// TIA Portal V21 export
// export: Created 2026-10-23T20:42:49.2153174Z, ExportSetting WithDefaults, DisplayName Totally Integrated Automation Portal, DisplayVersion V21 Update 1, DisplayName SINAMICS Startdrive Advanced, DisplayVersion V21 HF2, DisplayName SINAMICS Startdrive G110M, G120, G120C, G120D, G120P, G115D, DisplayVersion V21 HF2, DisplayName SINAMICS Startdrive G130, G150, S120, S150, G200, G220, S200, S210, S220, Innomotics MVD, DisplayVersion V21 HF2, DisplayName STEP 7 Professional, DisplayVersion V21 Update 1, DisplayName STEP 7 Safety, DisplayVersion V21, DisplayName Tech WebApplication, DisplayVersion V21, DisplayName WinCC Basic/Comfort/Advanced, DisplayVersion V21 Update 1, DisplayName WinCC Unified, DisplayVersion V21 Update 1
FUNCTION_BLOCK "FB_Mixed"   // FB9, LAD
TITLE = KOP-Baustein mit SCL-Netzwerk / LAD block with an SCL network
{ S7_Optimized_Access := 'TRUE' }
VERSION : 0.1
// stored: AutoNumber true, IsIECCheckEnabled false, IsRetainMemResEnabled false, MemoryReserve 100, SetENOAutomatically false, UDAEnableTagReadback false
   VAR_INPUT
      Start : Bool;   // Startbefehl / Start command
      RawValue : Int;   // Rohwert / Raw value
   END_VAR
   VAR_OUTPUT
      Running : Bool;   // Läuft / Running
      Scaled : Real;   // Skalierter Wert / Scaled value
      AboveLimit : Bool;   // Läuft und über dem Grenzwert / Running and above the limit
   END_VAR
   VAR
      Factor : Real := 2.5;   // Skalierungsfaktor / Scaling factor
      Limit : Real := 100.0;   // Grenzwert / Limit
      IsAbove : Bool;   // Skalierter Wert über dem Grenzwert / Scaled value above the limit
   END_VAR
BEGIN

REGION Network 1: KOP-Netzwerk vor dem SCL-Netzwerk / LAD network before the SCL network
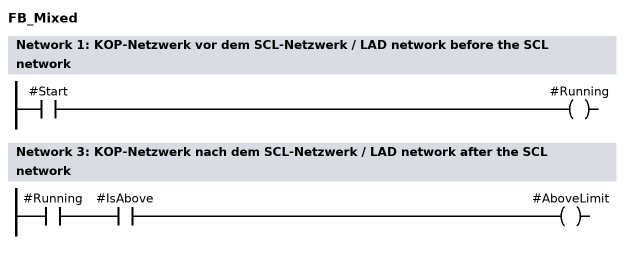
   RUNG wire#powerrail
      Contact( #Start )
      Coil( #Running )
   END_RUNG
   // the same network as SCL:
   #Running := #Start;
END_REGION

REGION Network 2 (SCL): SCL-Netzwerk im KOP-Baustein / SCL network inside the LAD block

       // Scale the raw value and compare it with the limit
       #Scaled := INT_TO_REAL(#RawValue) * #Factor;
       #IsAbove := #Scaled > #Limit;
END_REGION

REGION Network 3: KOP-Netzwerk nach dem SCL-Netzwerk / LAD network after the SCL network
   RUNG wire#powerrail
      Contact( #Running )
      Contact( #IsAbove )
      Coil( #AboveLimit )
   END_RUNG
   // the same network as SCL:
   #AboveLimit := #Running AND #IsAbove;
END_REGION
END_FUNCTION_BLOCK
